Fanuc KAREL source: KT00856.KL

PROGRAM KT00856
%NOLOCKGROUP
VAR
  I1: INTEGER
  I2: INTEGER
  OUT: INTEGER
BEGIN
  I1 = 2
  I2 = 3
  I1 = 2
  I2 = 3
  OUT = ROUND(I1)
END KT00856
